(* CODESYS project ciphersuite.library
   DefaultNamespace: KOSTAL.AF2024.Connectivity.TLS.CipherSuite.OpenSSL
   DocFormat: reStructuredText
   Description: Contains the cipher suites supported by Beckhoff in OpenSSL format.
   Author: Frank Dümpelmann
   Title: KOSTAL.AF2024.Connectivity.TLS.CipherSuite.OpenSSL
   Version: 1.0.0.0
   Company: KOSTAL GmbH & Co.KG
   Placeholder: KOSTAL.AF2024.Connectivity.TLS.CipherSuite.OpenSSL

Project tree, tasks and I/O mapping:
  Project Information/
    function F_GetCompany [ST]
    function F_GetTitle [ST]
    function F_GetVersion [ST]
  Version/
    global variables Global_Version
  global variables TLS_V1_2
*)

// Version/Global_Version
{attribute 'TcGenerated'}
{attribute 'no-analysis'}
{attribute 'linkalways'}
// This function has been automatically generated from the project information.
VAR_GLOBAL CONSTANT
	{attribute 'const_non_replaced'}
	stLibVersion_KOSTAL_AF2024_Connectivity_TLS_CipherSuite_OpenSSL : ST_LibVersion := (iMajor := 1, iMinor := 0, iBuild := 0, iRevision := 0, nFlags := 0, sVersion := '1.0.0.0');
END_VAR

// TLS_V1_2
{attribute 'qualified_only'}
VAR_GLOBAL CONSTANT
	
	DHE_RSA_AES256_SHA256		: STRING:='DHE-RSA-AES256-SHA256';
	ECDHE_RSA_AES256_SHA384	: STRING:='ECDHE-RSA-AES256-SHA384';
	ECDHE_ECDSA_AES256_SHA	: STRING:='ECDHE-ECDSA-AES256-SHA';
	ECDHE_RSA_AES256_SHA		: STRING:='ECDHE-RSA-AES256-SHA';
	DHE_RSA_AES256_SHA			: STRING:='DHE-RSA-AES256-SHA';
	ECDHE_ECDSA_AES128_GCM_SHA256	: STRING:='ECDHE-ECDSA-AES128-GCM-SHA256';
	ECDHE_RSA_AES128_GCM_SHA256	: STRING:='ECDHE-RSA-AES128-GCM-SHA256';
	DHE_RSA_AES128_GCM_SHA256	: STRING:='DHE-RSA-AES128-GCM-SHA256';
	ECDHE_ECDSA_AES128_SHA256: STRING:='ECDHE-ECDSA-AES128-SHA256';
	ECDHE_RSA_AES128_SHA256	: STRING:='ECDHE-RSA-AES128-SHA256';
	DHE_RSA_AES128_SHA256	: STRING:='DHE-RSA-AES128-SHA256';
	ECDHE_ECDSA_AES128_SHA	: STRING:='ECDHE-ECDSA-AES128-SHA';
	ECDHE_RSA_AES128_SHA	: STRING:='ECDHE-RSA-AES128-SHA';
	DHE_RSA_AES128_SHA	: STRING:='DHE-RSA-AES128-SHA';
	ECDHE_ECDSA_DES_CBC3_SHA	: STRING:='ECDHE-ECDSA-DES-CBC3-SHA';
	ECDHE_RSA_DES_CBC3_SHA	: STRING:='ECDHE-RSA-DES-CBC3-SHA';
	EDH_RSA_DES_CBC3_SHA	: STRING:='EDH-RSA-DES-CBC3-SHA';
	AES256_SHA256	: STRING:='AES256-SHA256';
	AES256_SHA	: STRING:='AES256-SHA';
	AES128_GCM_SHA256	: STRING:='AES128-GCM-SHA256';
	AES128_SHA256	: STRING:='AES128-SHA256';
	AES128_SHA	: STRING:='AES128-SHA';
	DES_CBC3_SHA	: STRING:='DES-CBC3-SHA';
	PSK_AES256_CBC_SHA	: STRING:='PSK-AES256-CBC-SHA';
	PSK_AES128_GCM_SHA256	: STRING:='PSK-AES128-GCM-SHA256';
	PSK_AES128_CBC_SHA256	: STRING:='PSK-AES128-CBC-SHA256';
	PSK_AES128_CBC_SHA	: STRING:='PSK-AES128-CBC-SHA';
	PSK_3DES_EDE_CBC_SHA	: STRING:='PSK-3DES-EDE-CBC-SHA';

END_VAR

// Project Information/F_GetCompany
// This function has been automatically generated from the project information.
{attribute 'signature_flag' := '1073741824'}
{attribute 'TcGenerated'}
{attribute 'no-analysis'}
FUNCTION F_GetCompany : WSTRING
VAR_INPUT
	
END_VAR

F_GetCompany := "KOSTAL GmbH & Co.KG";

END_FUNCTION

// Project Information/F_GetTitle
// This function has been automatically generated from the project information.
{attribute 'signature_flag' := '1073741824'}
{attribute 'TcGenerated'}
{attribute 'no-analysis'}
FUNCTION F_GetTitle : WSTRING
VAR_INPUT
	
END_VAR

F_GetTitle := "KOSTAL.AF2024.Connectivity.TLS.CipherSuite.OpenSSL";

END_FUNCTION

// Project Information/F_GetVersion
// This function has been automatically generated from the project information.
{attribute 'signature_flag' := '1073741824'}
{attribute 'TcGenerated'}
{attribute 'no-analysis'}
FUNCTION F_GetVersion : ST_LibVersion
VAR_INPUT
	
END_VAR

F_GetVersion.iMajor := 1;
F_GetVersion.iMinor := 0;
F_GetVersion.iBuild := 0;
F_GetVersion.iRevision := 0;
F_GetVersion.sVersion := '1.0.0.0';
F_GetVersion.nFlags := 0;

END_FUNCTION
